(* IEC 61131-3 sources: JingjiangArm/moonboxpro_arm_8.4/Application/Application/任务列表/TensionTask/张力控制/收放料/锥度控制, 11 files *)

(* ---- StPoint_XY.st ---- *)
(*@CES
Name=StPoint_XY
Type=Gvl
TypeGuid=2db5746d-d284-4425-9f7f-2663a34b0ebc
Guid=09f53c8f-47df-4e4e-acd6-e976559a9c39
HasDeclaration=True
HasImplementation=False
*)
{DECLARATION}
TYPE StPoint_XY :(*点位置-目前用于锥度(X=卷径|Y=气压)*)
STRUCT
	rX:REAL;
	rY:REAL;
END_STRUCT
END_TYPE

{IMPLEMENTATION}

(* ---- KS_CovertUnit_Taper.st ---- *)
(*@CES
Name=KS_CovertUnit_Taper
Type=FunctionBlock
TypeGuid=6f9dac99-8de1-4efc-8465-68ac443b7d08
Guid=64151f1e-8911-4786-9206-474c18fed1e9
HasDeclaration=True
HasImplementation=True
*)
{DECLARATION}
FUNCTION KS_CovertUnit_Taper : BOOL(*锥度单位转换|以%作为基准互相转换*)
(*如果参数出错了，则会重新处理单位变量|2022.10.16.104813*)
(*2025.1.15.152522 增加了停机张力值的处理@主要时针对收料*)
VAR_INPUT
	i_pbyUnit:POINTER TO BYTE;(*单位值|0-%|1-N|2-Mpa|参数非法按照百分比显示*)
	i_xConfirmN:BOOL;(*牛顿对应确认按钮*)
	i_xConfirmMpa:BOOL;(*Mpa对应确认按钮*)
	i_prConfirmTaperPercentMatchN:POINTER TO REAL;(*确认的百分比值-牛顿单位*)
	i_prConfirmTaperPercentMatchMpa:POINTER TO REAL;(*确认的百分比值-Mpa单位*)
	i_rConfirmTaperN: REAL;(*确认的牛顿值*)
	i_rConfirmTaperMpa: REAL;(*确认的Mpa值*)
	i_prTaperValueBegin_Hmi:POINTER TO REAL;(*界面锥度显示值-起始*)
	i_prTaperValueEnd_Hmi:POINTER TO REAL;(*界面锥度显示值-结束*)
	i_prTaperValueCur_Hmi:POINTER TO REAL;(*界面显示当前值|根据单位切换*)
	i_pbyLastUnit:POINTER TO BYTE;(*上个周期的单位选择值*)

	i_prTaperPencent_Begin:POINTER TO REAL;(*锥度起始百分比值*)
	i_prTaperPencent_End:POINTER TO REAL;(*锥度起始百分比值*)
	i_lrTaperPencent_Cur:LREAL;(*锥度起始百分比当前值*)

	(*2025.1.15.152522 增加了停机张力值的处理@主要时针对收料*)
	(*不用可以写0*)
	i_pbyInitTaper:POINTER TO BYTE;(*停机初始气压百分比*)
	i_prInitTaper_Hmi:POINTER TO REAL;(*收料初始气压显示值|根据单位切换*)

END_VAR
VAR
	lrConfirmTaperPencent: LREAL;(*确认的百分比值——和*)
	lrConfirmTaper: LREAL;(*确认的百分比对应的单位的值*)

	lrCoeff: LREAL;
END_VAR
{IMPLEMENTATION}
IF i_prConfirmTaperPercentMatchN<>0 AND
	i_prConfirmTaperPercentMatchMpa<>0 AND
	i_prTaperValueBegin_Hmi<>0 AND
	i_prTaperValueEnd_Hmi<>0 AND
	i_prTaperPencent_Begin<>0 AND
	i_pbyLastUnit<>0 AND
	i_pbyUnit<>0 AND
	i_prTaperValueCur_Hmi<>0 AND
	i_prTaperPencent_End<>0 THEN;
ELSE
	RETURN;
END_IF

(*确认对应关系|*)
IF i_xConfirmN THEN(*N确认|*)
	i_prConfirmTaperPercentMatchN^:=LREAL_TO_REAL(i_lrTaperPencent_Cur);
END_IF

IF i_xConfirmMpa THEN(*Mpa确认|*)
	i_prConfirmTaperPercentMatchMpa^:=LREAL_TO_REAL(i_lrTaperPencent_Cur);
END_IF

CASE i_pbyUnit^ OF
	1:(*单位N*)
		lrConfirmTaperPencent:=i_prConfirmTaperPercentMatchN^;
		lrConfirmTaper:=i_rConfirmTaperN;

		(*2022.10.16.104832 +*)
		IF lrConfirmTaperPencent=0 OR
			lrConfirmTaper=0 THEN
			i_pbyUnit^:=0;(*确认的系数出错了|不能切换单位*)
		END_IF
	2:(*单位Mpa*)
		lrConfirmTaperPencent:=i_prConfirmTaperPercentMatchMpa^;
		lrConfirmTaper:=i_rConfirmTaperMpa;
		(*2022.10.16.104832 +*)
		IF lrConfirmTaperPencent=0 OR
			lrConfirmTaper=0 THEN
			i_pbyUnit^:=0;(*确认的系数出错了|不能切换单位*)
		END_IF
ELSE(*单位%*)
	lrConfirmTaperPencent:=0;(*根据下面条件|使用百分比显示*)
	i_pbyUnit^:=0;
END_CASE

(*单位切换了|*)
lrCoeff:=1;
IF lrConfirmTaperPencent<>0 AND  lrConfirmTaper<>0 THEN
	lrCoeff:=(lrConfirmTaper)/lrConfirmTaperPencent;
END_IF

IF i_pbyLastUnit^ <> i_pbyUnit^ THEN(*将百分比值按照对应单位换算写入*)
	i_prTaperValueBegin_Hmi^:=LREAL_TO_REAL(lrCoeff*i_prTaperPencent_Begin^);
	i_prTaperValueEnd_Hmi^:=LREAL_TO_REAL(lrCoeff*i_prTaperPencent_End^);

	(*2025.1.15.152838+针对收料起始气压的处理输出*)
	IF i_prInitTaper_Hmi<>0 AND i_pbyInitTaper<>0 THEN
		i_prInitTaper_Hmi^:=LREAL_TO_REAL(lrCoeff*i_pbyInitTaper^);
	END_IF
ELSE
	i_prTaperPencent_Begin^:=LREAL_TO_REAL(i_prTaperValueBegin_Hmi^/lrCoeff);
	i_prTaperPencent_End^:=LREAL_TO_REAL(i_prTaperValueEnd_Hmi^/lrCoeff);
	(*最大100*)
	IF i_prTaperPencent_Begin^>100 THEN i_prTaperPencent_Begin^:=100;END_IF
	IF i_prTaperPencent_End^>100 THEN i_prTaperPencent_End^:=100;END_IF

	(*2025.1.15.152838+针对收料起始气压的处理输出*)
	IF i_prInitTaper_Hmi<>0 AND i_pbyInitTaper<>0 THEN
		i_pbyInitTaper^:=LREAL_TO_BYTE(i_prInitTaper_Hmi^/lrCoeff);
		IF i_pbyInitTaper^>100 THEN i_pbyInitTaper^:=100; END_IF
	END_IF

END_IF
(*当前值根据单位转换*)
i_prTaperValueCur_Hmi^:=LREAL_TO_REAL(lrCoeff*i_lrTaperPencent_Cur);
(*更新上个周期的单位值*)
i_pbyLastUnit^:=i_pbyUnit^;

(* ---- KS_GetCurveCoeff.st ---- *)
(*@CES
Name=KS_GetCurveCoeff
Type=FunctionBlock
TypeGuid=6f9dac99-8de1-4efc-8465-68ac443b7d08
Guid=9ebd4b66-811d-4a43-a8fd-0ccbf91fd938
HasDeclaration=True
HasImplementation=True
*)
{DECLARATION}
FUNCTION KS_GetCurveCoeff : BOOL(*锥度曲线拟合系数|支持直线和二次曲线*)
(*拟合系数-直线 Y=Ax+B
	   二次曲线 Y=Ax*x+Bx+C*)

(*支持多点计算(程序中允许100点输入)*)
(*-1 参数非法
  -2 直线拟合出错了*)
VAR_INPUT
	i_byCurveType:BYTE;(*曲线类型|=0 直线
								 |=1 二次曲线(点位太少按照直线输出)
								 |=2 三次曲线(暂不支持)*)
	i_iPoitNum_Max:INT;(*最大输入的点个数|根据这个值获取点位数据*)
	i_dwSaAdr_Point_XY:DWORD;(*点位数据的首地址|按照StPoint_XY结构体存放*)
	i_piValidPoitNum:POINTER TO INT;(*最大有效点个数*)
	(*拟合系数-直线 Y=Ax+B
		   二次曲线 Y=Ax*x+Bx+C*)
	i_prFitCoeff_A:POINTER TO REAL;(*拟合系数A*)
	i_prFitCoeff_B:POINTER TO REAL;(*拟合系数B*)
	i_prFitCoeff_C:POINTER TO REAL;(*拟合系数C*)
END_VAR
VAR
	in: INT;
	iPoitNum_Max: INT;(*最大点数*)
	astStPoint_XY:ARRAY [1..100] OF StPoint_XY;(*X轴为卷径|Y 为锥度值@按照100个点申请*)
	astValidStPoint_XY:ARRAY [1..100] OF StPoint_XY;(*X轴为卷径|Y 为锥度值@有效的点位*)
	iValidPoitNum:INT;(*有效点位的个数*)
	byCurveType: BYTE;(*曲线类型*)
	rA: REAL;
	rB: REAL;
	rC: REAL;
	xRtn: BOOL;
	iErrCode:INT;
END_VAR
{IMPLEMENTATION}
byCurveType:=i_byCurveType;
iPoitNum_Max:=i_iPoitNum_Max;
IF i_dwSaAdr_Point_XY<>0 THEN;
	SysMemCpy(ADR(astStPoint_XY),i_dwSaAdr_Point_XY,INT_TO_DWORD(iPoitNum_Max)*SIZEOF(astStPoint_XY[1]));
ELSE
	iErrCode:=-1;
END_IF

(*检查点位的合法性-X或者Y有一个=0认为是无效点*)
FOR iN:=1 TO iPoitNum_Max BY 1 DO
	IF astStPoint_XY[iN].rX=0 OR
		astStPoint_XY[iN].rY=0 THEN(*非法点，剔除*);
	ELSE
		iValidPoitNum:=iValidPoitNum+1;
		astValidStPoint_XY[iValidPoitNum]:=astStPoint_XY[iN];
	END_IF
END_FOR

(*曲线算法*)
byCurveType:=i_byCurveType;
CASE byCurveType OF
	0:(*直线拟合|*)
		xRtn:=KS_StraightLine(iValidPoitNum, ADR(astValidStPoint_XY), ADR(rA), ADR(rB));
		IF xRtn THEN
			iErrCode:=-2;
		END_IF
ELSE(*默认按照二次拟合*)
		xRtn:=KS_ParabolicLine(
					iValidPoitNum(*i_iValidPoitNum*),
					ADR(astValidStPoint_XY)(*i_pastValidStPoint_XY*),
					ADR(rA)(*i_prA*),
					ADR(rB)(*i_prB*),
					ADR(rC)(*i_prC*));
		IF xRtn THEN
			iErrCode:=-2;
		END_IF
END_CASE

IF i_piValidPoitNum<>0 THEN
	i_piValidPoitNum^:=iValidPoitNum;
END_IF
IF i_prFitCoeff_A<>0 THEN
	i_prFitCoeff_A^:=rA;
END_IF
IF i_prFitCoeff_B<>0 THEN
	i_prFitCoeff_B^:=rB;
END_IF

IF i_prFitCoeff_C<>0 THEN
	i_prFitCoeff_C^:=rC;
END_IF

KS_GetCurveCoeff:=iErrCode<>0;

(* ---- KS_ParabolicLine.st ---- *)
(*@CES
Name=KS_ParabolicLine
Type=FunctionBlock
TypeGuid=6f9dac99-8de1-4efc-8465-68ac443b7d08
Guid=32bb2783-1164-4a85-bd37-5e8616daa227
HasDeclaration=True
HasImplementation=True
*)
{DECLARATION}
FUNCTION KS_ParabolicLine : BOOL(*二次抛物线|Y=Ax^2+Bx+C@先不处理多点直线拟合|输出有效则报错*)
VAR_INPUT
	i_iValidPoitNum:INT;(*最大有效点个数*)
	i_pastValidStPoint_XY:POINTER TO ARRAY [1..100] OF StPoint_XY;(*X轴为卷径|Y 为锥度值@有效的点位*)
	i_prA:POINTER TO REAL;
	i_prB:POINTER TO REAL;
	i_prC:POINTER TO REAL;
END_VAR
VAR
	xParaErr:BOOL;
	arPoint_X:ARRAY [1..100] OF REAL;
	arPoint_Y:ARRAY [1..100] OF REAL;
	lrATemp:LREAL;
	lrBTemp:LREAL;
	rA:REAL;
	rB:REAL;
	rC:REAL;
	iN: INT;
	byType: BYTE;
	pstValidStPoint_XY:POINTER TO StPoint_XY;(*X轴为卷径|Y 为锥度值@有效的点位*)
	lrTemp: LREAL;
	lrTemp1: LREAL;
	lrTemp2: LREAL;
	lrTemp3: LREAL;
	lrTemp4: LREAL;
	lrTemp5: LREAL;
	lrTemp6: LREAL;
	lrTemp7: LREAL;
	lrAverage_X: LREAL;(*X的平均值*)
	lrAverage_Y: LREAL;(*Y的平均值*)
	lrAverage_XY: LREAL;(*XY的平均值*)
	lrAverage_X_Square2: LREAL;(*X^2的平均值*)
	lrAverage_X_Square3: LREAL;(*X^3的平均值*)
	lrAverage_X_Square4: LREAL;(*X^4的平均值*)
	lrAverage_XSquare2Y: LREAL;(*X^2*Y的平均值*)
END_VAR
{IMPLEMENTATION}
IF i_pastValidStPoint_XY<>0 THEN
	IF i_iValidPoitNum>=4 THEN(*4个点以上使用拟合算法*)
		byType:=3;
	ELSIF i_iValidPoitNum=3 THEN(*3个点使用抛物线*)
		byType:=2;
	ELSIF i_iValidPoitNum=2 THEN(*2个点使用直线*)
		byType:=1;
	ELSE(*点位太少*)
		xParaErr:=TRUE;
	END_IF

	IF NOT xParaErr THEN
		FOR iN:=1  TO i_iValidPoitNum BY 1 DO
			pstValidStPoint_XY:=ADR(i_pastValidStPoint_XY^[iN]);
			arPoint_X[iN]:=pstValidStPoint_XY^.rX;
			arPoint_Y[iN]:=pstValidStPoint_XY^.rY;
		END_FOR

		CASE byType OF
			1:(*直线*)
				lrTemp	:=arPoint_X[1]-arPoint_X[2];
				lrTemp1	:=arPoint_Y[1]-arPoint_Y[2];
				IF lrTemp<>0 THEN
					rA:=LREAL_TO_REAL(lrTemp1/lrTemp);

					lrTemp1:=arPoint_X[1]*arPoint_Y[2]-arPoint_X[2]*arPoint_Y[1];
					rB:=lrTemp1/lrTemp;
				ELSE
					xParaErr:=TRUE;
				END_IF

			2:(*抛物线*)
				(*计算rB*)
				lrTemp1:=(arPoint_X[2]*arPoint_X[2]-arPoint_X[3]*arPoint_X[3]);(*X2^2-X3^2*)
				lrTemp1:=lrTemp1*(arPoint_X[1]-arPoint_X[2]);(*lrTemp1*(X1-X2)*)
				lrTemp2:=(arPoint_X[1]*arPoint_X[1]-arPoint_X[2]*arPoint_X[2]);(*X1^2-X2^2*)
				lrTemp2:=lrTemp2*(arPoint_X[2]-arPoint_X[3]);(*lrTemp2*(X2-X3)*)
				lrTemp:=lrTemp1-lrTemp2;(*rB的分母*)

				IF lrTemp<>0 THEN
					lrTemp1:=(arPoint_X[2]*arPoint_X[2]-arPoint_X[3]*arPoint_X[3]);(*X2^2-X3^2*)
					lrTemp1:=lrTemp1*(arPoint_Y[1]-arPoint_Y[2]);(*lrTemp1*(Y1-Y2)*)
					lrTemp2:=(arPoint_X[1]*arPoint_X[1]-arPoint_X[2]*arPoint_X[2]);(*X1^2-X2^2*)
					lrTemp2:=lrTemp2*(arPoint_Y[2]-arPoint_Y[3]);(*lrTemp1*(Y2-Y3)*)

					rB:=(lrTemp1-lrTemp2)/lrTemp;
				ELSE
					xParaErr:=TRUE;
				END_IF

				(*计算rA*)
				IF NOT xParaErr THEN
					lrTemp:=(arPoint_X[1]*arPoint_X[1]-arPoint_X[2]*arPoint_X[2]);(*X1^2-X2^2*)
					IF lrTemp<>0 THEN
						lrTemp1:=arPoint_Y[1]-arPoint_Y[2]-rB*(arPoint_X[1]-arPoint_X[2]);(*Y1-Y2-rB*(X1-X2)*)
						rA:=lrTemp1/lrTemp;
					ELSE
						xParaErr:=TRUE;
					END_IF
				END_IF
				(*计算rC*)
				IF NOT xParaErr THEN
					rC:=arPoint_Y[1]-rA*(arPoint_X[1]*arPoint_X[1])-rB*arPoint_X[1];
				END_IF

			3:(*拟合曲线|*)
				lrTemp:=0;
				lrTemp1:=0;
				lrTemp2:=0;
				lrTemp3:=0;
				lrTemp4:=0;
				lrTemp5:=0;
				lrTemp6:=0;
				lrTemp7:=0;
				FOR iN:=1 TO i_iValidPoitNum BY 1 DO
					lrTemp1:=lrTemp1+arPoint_X[iN];
					lrTemp2:=lrTemp2+arPoint_Y[iN];
					lrTemp3:=lrTemp3+arPoint_X[iN]*arPoint_Y[iN];
					lrTemp4:=lrTemp4+arPoint_X[iN]*arPoint_X[iN];
					lrTemp5:=lrTemp5+arPoint_X[iN]*arPoint_X[iN]*arPoint_X[iN];
					lrTemp6:=lrTemp6+arPoint_X[iN]*arPoint_X[iN]*arPoint_X[iN]*arPoint_X[iN];
					lrTemp7:=lrTemp7+arPoint_X[iN]*arPoint_X[iN]*arPoint_Y[iN];
				END_FOR

				(*计算X Y的平均值*)
				lrAverage_X			:=lrTemp1/i_iValidPoitNum;
				lrAverage_Y			:=lrTemp2/i_iValidPoitNum;
				lrAverage_XY		:=lrTemp3/i_iValidPoitNum;
				lrAverage_X_Square2	:=lrTemp4/i_iValidPoitNum;
				lrAverage_X_Square3	:=lrTemp5/i_iValidPoitNum;
				lrAverage_X_Square4	:=lrTemp6/i_iValidPoitNum;
				lrAverage_XSquare2Y	:=lrTemp7/i_iValidPoitNum;

				(*计算拟合的rA*)
				lrTemp1:=lrAverage_X_Square3-lrAverage_X*lrAverage_X_Square2;
				lrTemp1:=lrTemp1*lrTemp1;
				lrTemp2:=lrAverage_X_Square4-lrAverage_X_Square2*lrAverage_X_Square2;
				lrTemp2:=lrTemp2*(lrAverage_X_Square2-lrAverage_X*lrAverage_X);
				lrTemp:=lrTemp1-lrTemp2;(*计算分母*)
				IF lrTemp<>0 THEN
					lrTemp1:=lrAverage_XY-lrAverage_X*lrAverage_Y;
					lrTemp1:=lrTemp1*(lrAverage_X_Square3-lrAverage_X*lrAverage_X_Square2);

					lrTemp2:=lrAverage_XSquare2Y-lrAverage_X_Square2*lrAverage_Y;
					lrTemp2:=lrTemp2*(lrAverage_X_Square2-lrAverage_X*lrAverage_X);
					lrATemp:=(lrTemp1-lrTemp2)/lrTemp;
					rA:=lrATemp;
				ELSE
					xParaErr:=TRUE;
				END_IF
				(*计算rB*)
				IF NOT xParaErr THEN
					lrTemp:=lrAverage_X_Square2-lrAverage_X*lrAverage_X;
					IF lrTemp<>0 THEN
						lrTemp1:=lrAverage_XY-lrAverage_X*lrAverage_Y-lrATemp*(lrAverage_X_Square3-lrAverage_X*lrAverage_X_Square2);
						lrBTemp:=lrTemp1/lrTemp;
						rB:=lrBTemp;
					ELSE
						xParaErr:=TRUE;
					END_IF
				END_IF

				(*计算rC*)
				IF NOT xParaErr THEN
					lrTemp:=lrAverage_Y-lrATemp*lrAverage_X_Square2-lrBTemp*lrAverage_X;
					rC:=lrTemp;
				END_IF
		ELSE;
		END_CASE

	END_IF
ELSE
	xParaErr:=TRUE;
END_IF

IF i_prA<>0 THEN
	i_prA^:=rA;
END_IF

IF i_prB<>0 THEN
	i_prB^:=rB;
END_IF

IF i_prC<>0 THEN
	i_prC^:=rC;
END_IF

KS_ParabolicLine:=xParaErr;

(* ---- KS_StraightLine.st ---- *)
(*@CES
Name=KS_StraightLine
Type=FunctionBlock
TypeGuid=6f9dac99-8de1-4efc-8465-68ac443b7d08
Guid=69642510-d218-426d-a290-8472573a37ba
HasDeclaration=True
HasImplementation=True
*)
{DECLARATION}
FUNCTION KS_StraightLine : BOOL(*直线|Y=Ax+B@先不处理多点直线拟合|输出有效则报错*)
VAR_INPUT
	i_iValidPoitNum:INT;(*最大有效点个数*)
	i_pastValidStPoint_XY:POINTER TO ARRAY [1..100] OF StPoint_XY;(*X轴为卷径|Y 为锥度值@有效的点位*)
	i_prA:POINTER TO REAL;
	i_prB:POINTER TO REAL;
END_VAR
VAR
	xParaErr:BOOL;
	arPoint_X:ARRAY [1..100] OF REAL;
	arPoint_Y:ARRAY [1..100] OF REAL;
	rA:REAL;
	rB:REAL;
	iN: INT;
	byType: BYTE;
	pstValidStPoint_XY:POINTER TO StPoint_XY;(*X轴为卷径|Y 为锥度值@有效的点位*)
	lrTemp: LREAL;
	lrTemp1: LREAL;
	lrTemp2: LREAL;
	lrTemp3: LREAL;
	lrTemp4: LREAL;
	lrSum_X: LREAL;
	lrSum_Y: LREAL;
	lrSum_XY: LREAL;
	lrSum_XSquart2: LREAL;
END_VAR
{IMPLEMENTATION}
IF i_pastValidStPoint_XY<>0 THEN
	IF i_iValidPoitNum>=3 THEN(*3个点以上使用拟合算法*)
		byType:=2;
	ELSIF i_iValidPoitNum=2 THEN(*2个点使用直线*)
		byType:=1;
	ELSE(*点位太少*)
		xParaErr:=TRUE;
	END_IF

	IF NOT xParaErr THEN
		FOR iN:=1  TO i_iValidPoitNum BY 1 DO
			pstValidStPoint_XY:=ADR(i_pastValidStPoint_XY^[iN]);
			arPoint_X[iN]:=pstValidStPoint_XY^.rX;
			arPoint_Y[iN]:=pstValidStPoint_XY^.rY;
		END_FOR

		CASE byType OF
			1:(*直线*)
				lrTemp	:=arPoint_X[1]-arPoint_X[2];
				lrTemp1	:=arPoint_Y[1]-arPoint_Y[2];
				IF lrTemp<>0 THEN
					rA:=LREAL_TO_REAL(lrTemp1/lrTemp);

					lrTemp1:=arPoint_X[1]*arPoint_Y[2]-arPoint_X[2]*arPoint_Y[1];
					rB:=LREAL_TO_REAL(lrTemp1/lrTemp);
				ELSE
					xParaErr:=TRUE;
				END_IF

			2:(*拟合直线*)
				lrSum_X:=0;
				lrSum_Y:=0;
				lrSum_XY:=0;
				lrSum_XSquart2:=0;
				FOR iN:=1 TO i_iValidPoitNum BY 1 DO
					lrSum_X:=lrSum_X+arPoint_X[iN];
					lrSum_Y:=lrSum_Y+arPoint_Y[iN];
					lrSum_XY:=lrSum_XY+arPoint_X[iN]*arPoint_Y[iN];
					lrSum_XSquart2:=lrSum_XSquart2+arPoint_X[iN]*arPoint_X[iN];
				END_FOR

				(*计算rB*)
				lrTemp:=i_iValidPoitNum*lrSum_XSquart2-lrSum_X*lrSum_X;
				IF lrTemp<>0 THEN
					lrTemp1:=lrSum_XSquart2*lrSum_Y-lrSum_X*lrSum_XY;
					rB:=LREAL_TO_REAL(lrTemp1/lrTemp);
				ELSE
					xParaErr:=TRUE;
				END_IF

				(*计算rA*)
				IF NOT xParaErr THEN
					lrTemp:=i_iValidPoitNum*lrSum_XSquart2-lrSum_X*lrSum_X;
					IF lrTemp<>0 THEN
						lrTemp1:=i_iValidPoitNum*lrSum_XY-lrSum_X*lrSum_Y;
						rA:=LREAL_TO_REAL(lrTemp1/lrTemp);
					ELSE
						xParaErr:=TRUE;
					END_IF
				END_IF
		ELSE;
		END_CASE

	END_IF
ELSE
	xParaErr:=TRUE;
END_IF

IF i_prA<>0 THEN
	i_prA^:=rA;
END_IF

IF i_prB<>0 THEN
	i_prB^:=rB;
END_IF

KS_StraightLine:=xParaErr;

(* ---- KS_Taper_Curve.st ---- *)
(*@CES
Name=KS_Taper_Curve
Type=FunctionBlock
TypeGuid=6f9dac99-8de1-4efc-8465-68ac443b7d08
Guid=9d8a75d4-e332-49bf-ad4d-ef60c80700c3
HasDeclaration=True
HasImplementation=True
*)
{DECLARATION}
FUNCTION KS_Taper_Curve : LREAL(*锥度1/X算法*)(*输出当前锥度*)
(*2025.1.9.162727  增加当前卷径输入*)
(*2025.2.26.163100 bug处理*)
VAR_INPUT
	i_rDiamCurAxis_Rw:REAL;(*2025.1.9.162744+*)
	i_rTaper_Begin_Rw: REAL;(*起始锥度*)
	i_rTaper_End_Rw: REAL;(*结束锥度*)
	i_rDiamTaper_Begin_Rw: REAL;(*起始锥度-直径*)
	i_rDiamTaper_End_Rw: REAL;(*结束锥度-直径*)
END_VAR
VAR
	lrMomentSa: LREAL;(*起始力矩*)
	lrMomentEd: LREAL;(*结束力矩*)
	lrCurrentMoment: LREAL;(*当前力矩*)
	lrCurrentTaper:LREAL;
END_VAR
{IMPLEMENTATION}
lrCurrentTaper:=0;
lrMomentSa:=(i_rTaper_Begin_Rw)*i_rDiamTaper_Begin_Rw;
lrMomentEd:=(i_rTaper_End_Rw)*i_rDiamTaper_End_Rw;

(*取消该限制@2025.2.26.163020*)
(*	IF lrMomentEd< lrMomentSa THEN lrMomentEd:=lrMomentSa;END_IF*)

IF i_rDiamCurAxis_Rw<= i_rDiamTaper_Begin_Rw THEN
	(*最小卷用最大张力*)
	lrCurrentTaper:= i_rTaper_Begin_Rw;
ELSIF i_rDiamCurAxis_Rw>= i_rDiamTaper_End_Rw THEN
	(*最大卷用最小张力*)
	lrCurrentTaper:= i_rTaper_End_Rw;
ELSE
	IF ( i_rDiamTaper_End_Rw-i_rDiamTaper_Begin_Rw)<>0 THEN
		lrCurrentMoment:=lrMomentSa+(lrMomentEd-lrMomentSa)*(i_rDiamCurAxis_Rw-i_rDiamTaper_Begin_Rw)
						/(i_rDiamTaper_End_Rw-i_rDiamTaper_Begin_Rw);
	ELSE
		lrCurrentMoment:=lrMomentSa;
	END_IF

	IF i_rDiamCurAxis_Rw<>0 THEN
		lrCurrentTaper:=lrCurrentMoment/i_rDiamCurAxis_Rw;
	ELSE
		lrCurrentTaper:=i_rTaper_Begin_Rw;
	END_IF
END_IF

KS_Taper_Curve:=lrCurrentTaper;

(* ---- KS_Taper_Straight.st ---- *)
(*@CES
Name=KS_Taper_Straight
Type=FunctionBlock
TypeGuid=6f9dac99-8de1-4efc-8465-68ac443b7d08
Guid=74716efb-2a9a-4cd3-af40-131a820a6ef5
HasDeclaration=True
HasImplementation=True
*)
{DECLARATION}
FUNCTION KS_Taper_Straight : LREAL(*锥度直线算法*)(*输出当前锥度*)
(*2025.1.9.162837 增加当前卷径输入*)
VAR_INPUT
	i_rDiamCurAxis_Rw:REAL;
	i_rTaper_Begin_Rw: REAL;(*起始锥度*)
	i_rTaper_End_Rw: REAL;(*结束锥度*)
	i_rDiamTaper_Begin_Rw: REAL;(*起始锥度-直径*)
	i_rDiamTaper_End_Rw: REAL;(*结束锥度-直径*)
END_VAR
VAR
	lrTempPercent: LREAL; (*临时用来计算%的变量*)
	lrCurrentTaper:LREAL;
END_VAR
{IMPLEMENTATION}
lrCurrentTaper:=0;
IF i_rDiamTaper_Begin_Rw<i_rDiamTaper_End_Rw THEN
	IF i_rDiamCurAxis_Rw<=i_rDiamTaper_Begin_Rw THEN
		(*最小卷用最大张力*)
		lrCurrentTaper:= i_rTaper_Begin_Rw;
	ELSIF i_rDiamCurAxis_Rw>=i_rDiamTaper_End_Rw THEN
		(*最大卷用最小张力*)
		lrCurrentTaper:= i_rTaper_End_Rw;
	ELSE
		(*卷径锥度的线性关系有效*)
		lrTempPercent:= (i_rDiamCurAxis_Rw - i_rDiamTaper_Begin_Rw) / (i_rDiamTaper_End_Rw - i_rDiamTaper_Begin_Rw);
		lrCurrentTaper:= i_rTaper_Begin_Rw - lrTempPercent * (i_rTaper_Begin_Rw - i_rTaper_End_Rw);
	END_IF
ELSE
	lrCurrentTaper:= 0;
END_IF
KS_Taper_Straight:=lrCurrentTaper;

(* ---- KS_FB_Taper.st ---- *)
(*@CES
Name=KS_FB_Taper
Type=FunctionBlock
TypeGuid=6f9dac99-8de1-4efc-8465-68ac443b7d08
Guid=684df15a-86b3-4c73-bdbe-f6eb8637542a
HasDeclaration=True
HasImplementation=True
*)
{DECLARATION}
FUNCTION_BLOCK KS_FB_Taper
(*2025.1.9.162926 增加了当前卷径输入接口@写到输入输出是为了防止漏改*)
(*2025.1.15.150823 停机锥度@防止停机张力投入时收料锥度设置过小引起的料膜被放料拉走问题*)
(*2025.3.7.112920 增加了多点直线和多点曲线的实现*)
(*2025.3.29.151033 停机锥度的实现更新丢了！麻烦*)
VAR_INPUT
	i_iGrpId: INT; (*1.A系;2.B系*)
	i_xTaperCurCTLEn:BOOL;(*当前锥度控制使能|在印刷状态且收牵合压或者色组至少合压一色时进行控制
						其他状态按照最大锥度输出|2021.8.30.164822*)
//	i_pstStShmGlobalParam: POINTER TO StShmGlobalParam; (*参数地址*)
	i_xTaperAdd:BOOL;
	i_xTaperDec:BOOL;
	i_rTaperMax:REAL;(*最大锥度限值值*)
	i_rTaperValue_Stop:REAL;(*停机锥度@防止停机张力投入时收料锥度设置过小引起的料膜被放料拉走问题*)

	i_byTaperAdjMode: BYTE;
	i_rDiamCurAxis: REAL;
	i_rTaper_Begin_Rw: REAL;(*起始锥度*)
	i_rTaper_End_Rw: REAL;(*结束锥度*)
	i_rDiamTaper_Begin_Rw: REAL;(*起始锥度-直径*)
	i_rDiamTaper_End_Rw: REAL;(*结束锥度-直径*)
END_VAR
VAR_OUTPUT
	o_rTaper_Cur: REAL;
END_VAR
VAR_IN_OUT
	iO_byTaperUnit: BYTE;
	io_rTaperValueBegin_Hmi: REAL;
	io_rTaperValueEnd_Hmi: REAL;
	io_astTaperPoint:ARRAY [1..10] OF StPoint_XY;
END_VAR
VAR
//	pstStGrpParam: POINTER TO StGrpParam; (*访问当前系参数的指针*)
	xTaperAdd:BOOL;
	xPreTaperAdd:BOOL;
	xTaperDec:BOOL;
	xPreTaperDec:BOOL;
	lrTemp: LREAL;
	lrCurrentTaper: LREAL;(*当前锥度值临时变量*)

	lrPreCurrentTaper: LREAL;(*上个周期的锥度*)
	lrDelTaper: LREAL;(*锥度的变化量*)
	iMaxTimeTOMaxTaper:INT:=200;(*到达最大锥度的周期次数，20ms周期时时间是4s*)
	iMaxTaper:INT:=100;(*最大锥度值*)

	(*2025.3.7.113256+byTaperAdjMode = 2*)
	xRtn: BOOL;
	iN: INT;
	iPoitMax: INT:=7;(*最大点数先按照7个*)
	iValidPoitNum: INT;(*实际有效的点数*)
	rFitCoeff_A: REAL;(*计算的二次系数*)
	rFitCoeff_B: REAL;(*计算的一次系数*)
	rFitCoeff_C: REAL;(*常量*)
	iMaxDiamIndex: INT;(*多点中卷径最大值索引*)
	iMinDiamIndex: INT;(*多点中卷径最小值索引*)
	rMinDiam: REAL;(*多点中最小卷径值*)
	rMaxDiam: REAL;(*多点中最大卷径值*)
END_VAR
{IMPLEMENTATION}
IF (i_iGrpId=1 OR i_iGrpId=2) THEN ;ELSE RETURN;END_IF

//pstStGrpParam:= ADR(i_pstStShmGlobalParam^.astStGrpParam[i_iGrpId]);

xTaperAdd:= i_xTaperAdd;
xTaperDec:= i_xTaperDec;

(*2022.2.23.112107 调整锥度界面加减逻辑*)
IF iO_byTaperUnit=1 THEN(*单位是N*)
	lrTemp:=1;
ELSIF iO_byTaperUnit=2 THEN(*单位是mpa*)
	lrTemp:=0.01;
ELSE(*单位是%*)
	lrTemp:=1;
END_IF

IF xTaperAdd AND NOT xPreTaperAdd THEN
	lrTemp:=lrTemp;
ELSIF xTaperDec AND NOT xPreTaperDec THEN
	lrTemp:=-lrTemp;
ELSE
	lrTemp:=0;
END_IF
(*
pstStGrpParam^.lrTaper_Begin_Rw:= pstStGrpParam^.lrTaper_Begin_Rw+lrTemp;
pstStGrpParam^.lrTaper_End_Rw:= pstStGrpParam^.lrTaper_End_Rw+lrTemp;
*)
(*2022.2.23.112206 处理的变量修改为带hmi界面的*)

io_rTaperValueBegin_Hmi:= io_rTaperValueBegin_Hmi+lrTemp;
io_rTaperValueEnd_Hmi:= io_rTaperValueEnd_Hmi+lrTemp;

IF 	io_rTaperValueBegin_Hmi>i_rTaperMax THEN
	io_rTaperValueBegin_Hmi:= i_rTaperMax;
ELSIF io_rTaperValueBegin_Hmi<0 THEN
	io_rTaperValueBegin_Hmi:=0;
END_IF

IF 	io_rTaperValueEnd_Hmi>i_rTaperMax THEN
	io_rTaperValueEnd_Hmi:= i_rTaperMax;
ELSIF io_rTaperValueEnd_Hmi<0 THEN
	io_rTaperValueEnd_Hmi:=0;
END_IF

xPreTaperAdd:=xTaperAdd;
xPreTaperDec:=xTaperDec;

(*
(*2019.4.11.164149 将锥度控制移植到功能块中.并额外增加了新的算法*)
CASE i_pstStShmGlobalParam^.stStSystemExtInfo.byTaperAdjMode OF
1:
	lrCurrentTaper:=KS_Taper_Curve(pstStGrpParam^.lrDiamCurAxis_Rw,pstStGrpParam);
ELSE
	lrCurrentTaper:=KS_Taper_Straight(pstStGrpParam^.lrDiamCurAxis_Rw,pstStGrpParam);
END_CASE

(*2021.8.30.164530 |*)
(*不控制的时候按照最大锥度输出*)
IF NOT i_xTaperCurCTLEn THEN
	lrCurrentTaper:=MAX(pstStGrpParam^.lrTaper_Begin_Rw,pstStGrpParam^.lrTaper_End_Rw);(*取最大值*)
	(*增加一个变量单独控制停机的锥度*)
	lrCurrentTaper:=MAX(lrCurrentTaper,i_rTaperValue_Stop);
END_IF
*)

(*2025.3.7.112958 +*)
(*2019.4.11.164149 将锥度控制移植到功能块中.并额外增加了新的算法*)
(*0--2变化*)
xRtn:=FALSE;
CASE i_byTaperAdjMode OF
1:(*2点曲线*)

	lrCurrentTaper:=KS_Taper_Curve(
			i_rDiamCurAxis,
			i_rTaper_Begin_Rw,
			i_rTaper_End_Rw,
			i_rDiamTaper_Begin_Rw,
			i_rDiamTaper_End_Rw
			);

	(*2021.8.30.164530 |*)
	(*不控制的时候按照最大锥度输出*)
	IF NOT i_xTaperCurCTLEn THEN
(*
		lrCurrentTaper:=MAX(pstStGrpParam^.lrTaper_Begin_Rw,pstStGrpParam^.lrTaper_End_Rw);(*取最大值*)
		(*增加一个变量单独控制停机的锥度*)
		lrCurrentTaper:=MAX(lrCurrentTaper,i_rTaperValue_Stop);
*)
		(*2025.3.29.151947+*)
		lrCurrentTaper:=i_rTaperValue_Stop;
	END_IF

2:(*多点曲线@2025.2.28.235627+*)
	(*寻找卷径锥度的最大值和最小值@限制输出使用*)
	iMinDiamIndex:=0;
	iMaxDiamIndex:=0;
	FOR iN:=1 TO iPoitMax BY 1 DO
		(*最小卷径值的索引*)
		IF iMinDiamIndex=0 THEN(*先找起始索引*)
			IF io_astTaperPoint[iN].rX<>0 THEN
				iMinDiamIndex:=iN;
			END_IF
		ELSE(*找到了第一个值*)
			IF io_astTaperPoint[iN].rX < io_astTaperPoint[iMinDiamIndex].rX THEN
				iMinDiamIndex:=iN;(*更新索引值*)
			END_IF
		END_IF

		(*最大卷径的索引*)
		IF iMaxDiamIndex=0 THEN(*先找起始索引*)
			IF io_astTaperPoint[iN].rX<>0 THEN
				iMaxDiamIndex:=iN;
			END_IF
		ELSE(*找到了第一个值*)
			IF io_astTaperPoint[iN].rX > io_astTaperPoint[iMaxDiamIndex].rX THEN
				iMaxDiamIndex:=iN;(*更新索引值*)
			END_IF
		END_IF
	END_FOR

	xRtn:=KS_GetCurveCoeff(
			1(*i_byCurveType*),
			iPoitMax(*i_iPoitNum_Max*),
			ADR(io_astTaperPoint[1])(*i_dwSaAdr_Point_XY*),
			ADR(iValidPoitNum)(*i_piValidPoitNum*),
			ADR(rFitCoeff_A)(*i_prFitCoeff_A*),
			ADR(rFitCoeff_B)(*i_prFitCoeff_B*),
			ADR(rFitCoeff_C)(*i_prFitCoeff_C*));
	(*输出的形式是a*x*x+b*x+C*)
	IF NOT xRtn THEN(*未报错@至少2个点*)
		lrCurrentTaper:=rFitCoeff_A*i_rDiamCurAxis*i_rDiamCurAxis+
						rFitCoeff_B*i_rDiamCurAxis+
						rFitCoeff_C;
		(*限值处理*)
		IF	iMinDiamIndex>0 AND iMinDiamIndex<=iPoitMax AND(*索引合法判断*)
			iMaxDiamIndex>0 AND iMaxDiamIndex<=iPoitMax THEN(*索引合法判断*)
			(*最小值处理*)
			rMinDiam:= io_astTaperPoint[iMinDiamIndex].rX;
			IF i_rDiamCurAxis<=rMinDiam THEN
				lrCurrentTaper:=rFitCoeff_A*rMinDiam*rMinDiam+
								rFitCoeff_B*rMinDiam+
								rFitCoeff_C;
			END_IF
			(*最大值处理*)
			rMaxDiam:= io_astTaperPoint[iMaxDiamIndex].rX;
			IF i_rDiamCurAxis>=rMaxDiam THEN
				lrCurrentTaper:=rFitCoeff_A*rMaxDiam*rMaxDiam+
								rFitCoeff_B*rMaxDiam+
								rFitCoeff_C;
			END_IF
(*
			(*2025.3.3.112928 调整*)
			(*2021.8.30.164530 |*)
			(*不控制的时候按照最大锥度输出*)
			IF NOT i_xTaperCurCTLEn THEN
				lrCurrentTaper:=MAX(rFitCoeff_A*rMinDiam*rMinDiam+rFitCoeff_B*rMinDiam+rFitCoeff_C,
								rFitCoeff_A*rMaxDiam*rMaxDiam+rFitCoeff_B*rMaxDiam+rFitCoeff_C);(*取最大值*)
				(*增加一个变量单独控制停机的锥度*)
				lrCurrentTaper:=MAX(lrCurrentTaper,i_rTaperValue_Stop);

			END_IF
*)
		ELSE
			lrCurrentTaper:=22.2;(*就随便给一个特殊值吧@有可能能指导查找问题*)
		END_IF
	ELSE(*拟合失败了@按照最大点输出*)
		IF iMaxDiamIndex>0 AND iMaxDiamIndex<=iPoitMax THEN(*索引合法判断*)
			lrCurrentTaper:=io_astTaperPoint[iMaxDiamIndex].rY;
		END_IF
	END_IF

	(*2025.3.29.151918+*)
	(*不控制的时候按照最大锥度输出*)
	IF NOT i_xTaperCurCTLEn THEN
		lrCurrentTaper:=i_rTaperValue_Stop;
	END_IF
ELSE(*2点直线*)
	lrCurrentTaper:=KS_Taper_Straight(
			i_rDiamCurAxis,
			i_rTaper_Begin_Rw,
			i_rTaper_End_Rw,
			i_rDiamTaper_Begin_Rw,
			i_rDiamTaper_End_Rw
			);

	(*2021.8.30.164530 |*)
	(*不控制的时候按照最大锥度输出*)
	IF NOT i_xTaperCurCTLEn THEN
(*
		lrCurrentTaper:=MAX(pstStGrpParam^.lrTaper_Begin_Rw,pstStGrpParam^.lrTaper_End_Rw);(*取最大值*)
		(*增加一个变量单独控制停机的锥度*)
		lrCurrentTaper:=MAX(lrCurrentTaper,i_rTaperValue_Stop);
*)
		(*2025.3.29.151937+*)
		lrCurrentTaper:=i_rTaperValue_Stop;
	END_IF
END_CASE

lrDelTaper:=INT_TO_LREAL(iMaxTaper)/INT_TO_LREAL(iMaxTimeTOMaxTaper);
(*rWatch:=lrCurrentTaper;*)
IF lrCurrentTaper> lrPreCurrentTaper THEN
	IF (lrCurrentTaper-lrPreCurrentTaper) > lrDelTaper THEN
		lrCurrentTaper:=lrPreCurrentTaper+lrDelTaper;
	ELSE;
	END_IF
ELSIF  lrCurrentTaper< lrPreCurrentTaper THEN
	IF (lrPreCurrentTaper-lrCurrentTaper) > lrDelTaper THEN
		lrCurrentTaper:=lrPreCurrentTaper-lrDelTaper;
	ELSE;
	END_IF
ELSE;
END_IF

o_rTaper_Cur:= LREAL_TO_REAL(lrCurrentTaper);
lrPreCurrentTaper:=lrCurrentTaper;

(* ---- KS_FB_Taper_UwRw_IfOf.st ---- *)
(*@CES
Name=KS_FB_Taper_UwRw_IfOf
Type=FunctionBlock
TypeGuid=6f9dac99-8de1-4efc-8465-68ac443b7d08
Guid=4508f757-99f8-49ac-966d-1f120aaadfc2
HasDeclaration=True
HasImplementation=True
*)
{DECLARATION}
FUNCTION_BLOCK KS_FB_Taper_UwRw_IfOf
VAR_INPUT
	i_xEn: BOOL;
END_VAR
VAR_OUTPUT
END_VAR
VAR
	fbKS_FB_TaperUnitDeal: KS_FB_TaperUnitDeal;
	(*锥度变化临时变量|只处理放料 放牵收牵*)
	rMaxTaper:REAL:=100;(*最大锥度|目前使用%*)
	iTimeTaperChange:INT:=10000;(*锥度变化时间|ms*)
	rTaperTar: REAL;
	rTaperCur: REAL;
	rDeltTaper: REAL;
	xInit_Taper_Cur: BOOL;
END_VAR
{IMPLEMENTATION}
IF i_xEn THEN
	(*2021.7.29.094016 张力单位切换控制逻辑|以及标定逻辑*)
	fbKS_FB_TaperUnitDeal(i_pstStGrpParam:=pstStGrpParam );

	(*处理4个锥度|放料、放牵、收料、收牵*)
	(*需要确定是否需要进行单位转换|目前是%*)
	(*使用起始锥度作为界面显示|当前锥度做规划*)
	(*放料*)
	(*由于当前锥度是保持型的|在这里做开机初始复位处理|*)
	IF NOT xInit_Taper_Cur THEN
		xInit_Taper_Cur:=TRUE;
		pstStGrpParam^.lrTaper_Cur_Uw:=0;
		pstStGrpParam^.lrTaper_Cur_If:=0;
		pstStGrpParam^.lrTaper_Cur_Of:=0;
	END_IF

	rTaperTar:=pstStGrpParam^.lrTaper_Begin_Uw;
	rTaperCur:=pstStGrpParam^.lrTaper_Cur_Uw;
	rDeltTaper:=rMaxTaper/iTimeTaperChange*gc_iCycleTime_Plc;
	IF rTaperCur<rTaperTar THEN
		rTaperCur:=rTaperCur+rDeltTaper;
		IF rTaperCur>=rTaperTar THEN
			rTaperCur:=rTaperTar;
		END_IF
	ELSIF rTaperCur>rTaperTar THEN
		rTaperCur:=rTaperCur-rDeltTaper;
		IF rTaperCur<=rTaperTar THEN
			rTaperCur:=rTaperTar;
		END_IF
	ELSE;
	END_IF
	pstStGrpParam^.lrTaper_Cur_Uw:=rTaperCur;
	(*放牵*)
	rTaperTar:=pstStGrpParam^.lrTaper_Begin_If;
	rTaperCur:=pstStGrpParam^.lrTaper_Cur_If;
	rDeltTaper:=rMaxTaper/iTimeTaperChange*gc_iCycleTime_Plc;
	IF rTaperCur<rTaperTar THEN
		rTaperCur:=rTaperCur+rDeltTaper;
		IF rTaperCur>=rTaperTar THEN
			rTaperCur:=rTaperTar;
		END_IF
	ELSIF rTaperCur>rTaperTar THEN
		rTaperCur:=rTaperCur-rDeltTaper;
		IF rTaperCur<=rTaperTar THEN
			rTaperCur:=rTaperTar;
		END_IF
	ELSE;
	END_IF
	pstStGrpParam^.lrTaper_Cur_If:=rTaperCur;
	(*收牵*)
	rTaperTar:=pstStGrpParam^.lrTaper_Begin_Of;
	rTaperCur:=pstStGrpParam^.lrTaper_Cur_Of;
	rDeltTaper:=rMaxTaper/iTimeTaperChange*gc_iCycleTime_Plc;
	IF rTaperCur<rTaperTar THEN
		rTaperCur:=rTaperCur+rDeltTaper;
		IF rTaperCur>=rTaperTar THEN
			rTaperCur:=rTaperTar;
		END_IF
	ELSIF rTaperCur>rTaperTar THEN
		rTaperCur:=rTaperCur-rDeltTaper;
		IF rTaperCur<=rTaperTar THEN
			rTaperCur:=rTaperTar;
		END_IF
	ELSE;
	END_IF
	pstStGrpParam^.lrTaper_Cur_Of:=rTaperCur;
END_IF

(* ---- KS_FB_TaperUnitDeal.st ---- *)
(*@CES
Name=KS_FB_TaperUnitDeal
Type=FunctionBlock
TypeGuid=6f9dac99-8de1-4efc-8465-68ac443b7d08
Guid=440da615-589b-45d5-ab61-0644875fc808
HasDeclaration=True
HasImplementation=True
*)
{DECLARATION}
FUNCTION_BLOCK KS_FB_TaperUnitDeal(*锥度单位处理*)
(*调整不同单位张力最大值的切换代码执行位置|2022.10.16.105041*)
(*2025.1.15.152035 计算收料停机锥度显示值*)
VAR_INPUT
	i_xEn: BOOL;
END_VAR
VAR_OUTPUT
END_VAR
VAR_IN_OUT
	io_byTaperUnitType:BYTE;(*张力单位切换标志|.0 放牵\.1收牵\.2放料\.3收料*)
	io_byTaperUnit_If: BYTE;
	io_byTaperUnit_Of: BYTE;
	io_byTaperUnit_Uw: BYTE;
	io_byTaperUnit_Rw: BYTE;
	io_byTaperUnitConfirm_Uw : BYTE;

END_VAR
VAR
	byLastUnit_Uw: BYTE:=3;(*初始化给一个不一样的值|用于触发开机取初值*)
	byLastUnit_Rw: BYTE:=3;(*初始化给一个不一样的值|用于触发开机取初值*)
	byLastUnit_If: BYTE:=3;(*初始化给一个不一样的值|用于触发开机取初值*)
	byLastUnit_Of: BYTE:=3;(*初始化给一个不一样的值|用于触发开机取初值*)
END_VAR
{IMPLEMENTATION}
IF i_xEn THEN;
ELSE
	RETURN;
END_IF

(**处理单位切换标志*)
IF io_byTaperUnitType<>0 THEN
	IF io_byTaperUnitType.0 THEN(*放牵切换*)
		io_byTaperUnit_If:=io_byTaperUnit_If+1;
		IF io_byTaperUnit_If>2 THEN
			io_byTaperUnit_If:=0;
		END_IF
	ELSIF io_byTaperUnitType.1 THEN(*收牵切换*)
		io_byTaperUnit_Of:=io_byTaperUnit_Of+1;
		IF io_byTaperUnit_Of>2 THEN
			io_byTaperUnit_Of:=0;
		END_IF
	ELSIF io_byTaperUnitType.2 THEN(*放料切换*)
		io_byTaperUnit_Uw:=io_byTaperUnit_Uw+1;
		IF io_byTaperUnit_Uw>2 THEN
			io_byTaperUnit_Uw:=0;
		END_IF
	ELSIF io_byTaperUnitType.3 THEN(*收料切换*)
		io_byTaperUnit_Rw:=io_byTaperUnit_Rw+1;
		IF io_byTaperUnit_Rw>2 THEN
			io_byTaperUnit_Rw:=0;
		END_IF
	ELSE;
	END_IF
	(*清除单位切换按钮*)
	io_byTaperUnitType:=0;
END_IF

(*放料处理*)
(*
g_rTaperMax_Uw:=100;
IF io_byTaperUnit_Uw=1 THEN(*放料单位|N*)
	g_rTaperMax_Uw:=500;
ELSIF io_byTaperUnit_Uw=2 THEN(*放料单位|Mpa*)
	g_rTaperMax_Uw:=1;
END_IF
*)
KS_CovertUnit_Taper(
	ADR(io_byTaperUnit_Uw)(*i_pbyUnit*),
	i_pstStGrpParam^.byTaperUnitConfirm_Uw.0(*i_xConfirmN*),
	i_pstStGrpParam^.byTaperUnitConfirm_Uw.1(*i_xConfirmMpa*),
	ADR(i_pstStGrpParam^.rPercentMatchN_Uw)(*i_prConfirmTaperPercentMatchN*),
	ADR(i_pstStGrpParam^.rPercentMatchMpa_Uw)(*i_prConfirmTaperPercentMatchMpa*),
	i_pstStGrpParam^.rN_Uw(*i_rConfirmTaperN*),
	i_pstStGrpParam^.rMpa_Uw(*i_rConfirmTaperMpa*),
	ADR(i_pstStGrpParam^.rTaperValueBegin_Hmi_Uw)(*i_prTaperValueBegin_Hmi*),
	ADR(i_pstStGrpParam^.rTaperValueEnd_Hmi_Uw)(*i_prTaperValueEnd_Hmi*),
	ADR(i_pstStGrpParam^.rTaperValueCur_Hmi_Uw)(*i_prTaperValueCur_Hmi*),

	ADR(byLastUnit_Uw)(*i_pbyLastUnit*),
	ADR(i_pstStGrpParam^.lrTaper_Begin_Uw)(*i_plrTaperPencent_Begin*),
	ADR(i_pstStGrpParam^.lrTaper_End_Uw)(*i_plrTaperPencent_End*),
	i_pstStGrpParam^.lrTaper_Cur_Uw(*i_lrTaperPencent_Cur*),
	(*2025.1.15.153326+*)
	0(*i_pbyInitTaper*),
	0(*i_prInitTaper_Hmi*));
(*2022.10.16.104937*)
g_rTaperMax_Uw:=100;
IF io_byTaperUnit_Uw=1 THEN(*放料单位|N*)
	g_rTaperMax_Uw:=500;
ELSIF io_byTaperUnit_Uw=2 THEN(*放料单位|Mpa*)
	g_rTaperMax_Uw:=1;
END_IF
(*清除确认按钮*)
i_pstStGrpParam^.byTaperUnitConfirm_Uw:=0;

(*收料处理*)
(*
g_rTaperMax_Rw:=100;
IF io_byTaperUnit_Rw=1 THEN(*放料单位|N*)
	g_rTaperMax_Rw:=500;
ELSIF io_byTaperUnit_Rw=2 THEN(*放料单位|Mpa*)
	g_rTaperMax_Rw:=1;
END_IF
*)
KS_CovertUnit_Taper(
	ADR(io_byTaperUnit_Rw)(*i_pbyUnit*),
	i_pstStGrpParam^.byTaperUnitConfirm_Rw.0(*i_xConfirmN*),
	i_pstStGrpParam^.byTaperUnitConfirm_Rw.1(*i_xConfirmMpa*),
	ADR(i_pstStGrpParam^.rPercentMatchN_Rw)(*i_prConfirmTaperPercentMatchN*),
	ADR(i_pstStGrpParam^.rPercentMatchMpa_Rw)(*i_prConfirmTaperPercentMatchMpa*),
	i_pstStGrpParam^.rN_Rw(*i_rConfirmTaperN*),
	i_pstStGrpParam^.rMpa_Rw(*i_rConfirmTaperMpa*),
	ADR(i_pstStGrpParam^.rTaperValueBegin_Hmi_Rw)(*i_prTaperValueBegin_Hmi*),
	ADR(i_pstStGrpParam^.rTaperValueEnd_Hmi_Rw)(*i_prTaperValueEnd_Hmi*),
	ADR(i_pstStGrpParam^.rTaperValueCur_Hmi_Rw)(*i_prTaperValueCur_Hmi*),
	ADR(byLastUnit_Rw)(*i_pbyLastUnit*),
	ADR(i_pstStGrpParam^.lrTaper_Begin_Rw)(*i_plrTaperPencent_Begin*),
	ADR(i_pstStGrpParam^.lrTaper_End_Rw)(*i_plrTaperPencent_End*),
	i_pstStGrpParam^.lrTaper_Cur_Rw(*i_lrTaperPencent_Cur*),
	(*2025.1.15.153326+*)
	ADR(i_pstStGrpParam^.byInitTaper_Rw)(*i_pbyInitTaper*),
	ADR(i_pstStGrpParam^.rInitTaper_Hmi_Rw)(*i_prInitTaper_Hmi*));
(*2022.10.16.104955*)
g_rTaperMax_Rw:=100;
IF io_byTaperUnit_Rw=1 THEN(*放料单位|N*)
	g_rTaperMax_Rw:=500;
ELSIF io_byTaperUnit_Rw=2 THEN(*放料单位|Mpa*)
	g_rTaperMax_Rw:=1;
END_IF
(*清除确认按钮*)
i_pstStGrpParam^.byTaperUnitConfirm_Rw:=0;

(*放牵处理*)
(*
g_rTaperMax_If:=100;
IF io_byTaperUnit_If=1 THEN(*放料单位|N*)
	g_rTaperMax_If:=500;
ELSIF io_byTaperUnit_If=2 THEN(*放料单位|Mpa*)
	g_rTaperMax_If:=1;
END_IF
*)
KS_CovertUnit_Taper(
	ADR(io_byTaperUnit_If)(*i_pbyUnit*),
	i_pstStGrpParam^.byTaperUnitConfirm_If.0(*i_xConfirmN*),
	i_pstStGrpParam^.byTaperUnitConfirm_If.1(*i_xConfirmMpa*),
	ADR(i_pstStGrpParam^.rPercentMatchN_If)(*i_prConfirmTaperPercentMatchN*),
	ADR(i_pstStGrpParam^.rPercentMatchMpa_If)(*i_prConfirmTaperPercentMatchMpa*),
	i_pstStGrpParam^.rN_If(*i_rConfirmTaperN*),
	i_pstStGrpParam^.rMpa_If(*i_rConfirmTaperMpa*),
	ADR(i_pstStGrpParam^.rTaperValueBegin_Hmi_If)(*i_prTaperValueBegin_Hmi*),
	ADR(i_pstStGrpParam^.rTaperValueEnd_Hmi_If)(*i_prTaperValueEnd_Hmi*),
	ADR(i_pstStGrpParam^.rTaperValueCur_Hmi_If)(*i_prTaperValueCur_Hmi*),
	ADR(byLastUnit_If)(*i_pbyLastUnit*),
	ADR(i_pstStGrpParam^.lrTaper_Begin_If)(*i_plrTaperPencent_Begin*),
	ADR(i_pstStGrpParam^.lrTaper_End_If)(*i_plrTaperPencent_End*),
	i_pstStGrpParam^.lrTaper_Cur_If(*i_lrTaperPencent_Cur*),
	(*2025.1.15.153326+*)
	0(*i_pbyInitTaper*),
	0(*i_prInitTaper_Hmi*));
(*2022.10.16.105013*)
g_rTaperMax_If:=100;
IF io_byTaperUnit_If=1 THEN(*放料单位|N*)
	g_rTaperMax_If:=500;
ELSIF io_byTaperUnit_If=2 THEN(*放料单位|Mpa*)
	g_rTaperMax_If:=1;
END_IF
(*清除确认按钮*)
i_pstStGrpParam^.byTaperUnitConfirm_If:=0;

(*收牵处理*)
(*
g_rTaperMax_of:=100;
IF io_byTaperUnit_Of=1 THEN(*放料单位|N*)
	g_rTaperMax_of:=500;
ELSIF io_byTaperUnit_Of=2 THEN(*放料单位|Mpa*)
	g_rTaperMax_of:=1;
END_IF
*)
KS_CovertUnit_Taper(
	ADR(io_byTaperUnit_Of)(*i_pbyUnit*),
	i_pstStGrpParam^.byTaperUnitConfirm_Of.0(*i_xConfirmN*),
	i_pstStGrpParam^.byTaperUnitConfirm_Of.1(*i_xConfirmMpa*),
	ADR(i_pstStGrpParam^.rPercentMatchN_Of)(*i_prConfirmTaperPercentMatchN*),
	ADR(i_pstStGrpParam^.rPercentMatchMpa_Of)(*i_prConfirmTaperPercentMatchMpa*),
	i_pstStGrpParam^.rN_Of(*i_rConfirmTaperN*),
	i_pstStGrpParam^.rMpa_Of(*i_rConfirmTaperMpa*),
	ADR(i_pstStGrpParam^.rTaperValueBegin_Hmi_Of)(*i_prTaperValueBegin_Hmi*),
	ADR(i_pstStGrpParam^.rTaperValueEnd_Hmi_Of)(*i_prTaperValueEnd_Hmi*),
	ADR(i_pstStGrpParam^.rTaperValueCur_Hmi_Of)(*i_prTaperValueCur_Hmi*),
	ADR(byLastUnit_Of)(*i_pbyLastUnit*),
	ADR(i_pstStGrpParam^.lrTaper_Begin_Of)(*i_plrTaperPencent_Begin*),
	ADR(i_pstStGrpParam^.lrTaper_End_Of)(*i_plrTaperPencent_End*),
	i_pstStGrpParam^.lrTaper_Cur_Of(*i_lrTaperPencent_Cur*),
	(*2025.1.15.153326+*)
	0(*i_pbyInitTaper*),
	0(*i_prInitTaper_Hmi*));
(*2022.10.16.105028*)
g_rTaperMax_of:=100;
IF io_byTaperUnit_Of=1 THEN(*放料单位|N*)
	g_rTaperMax_of:=500;
ELSIF io_byTaperUnit_Of=2 THEN(*放料单位|Mpa*)
	g_rTaperMax_of:=1;
END_IF
(*清除确认按钮*)
i_pstStGrpParam^.byTaperUnitConfirm_Of:=0;

(* ---- KS_FB_TaperUnitDeal_New.st ---- *)
(*@CES
Name=KS_FB_TaperUnitDeal_New
Type=FunctionBlock
TypeGuid=6f9dac99-8de1-4efc-8465-68ac443b7d08
Guid=029751e0-fe3d-4f68-a3f4-ab7fe94fc43b
HasDeclaration=True
HasImplementation=True
*)
{DECLARATION}
FUNCTION_BLOCK KS_FB_TaperUnitDeal_New(*锥度单位处理*)
(*调整不同单位张力最大值的切换代码执行位置|2022.10.16.105041*)
(*2025.1.15.152035 计算收料停机锥度显示值*)
VAR_INPUT
	i_xEn: BOOL;
	i_rN: REAL;
	i_rMpa: REAL;
	i_pbyInitTaper: POINTER TO BYTE;
	i_prInitTaper_Hmi: POINTER TO REAL;
END_VAR
VAR_OUTPUT
END_VAR
VAR_IN_OUT
	io_xTaperUnitType:BOOL;(*张力单位切换标志|.0 放牵\.1收牵\.2放料\.3收料*)
	io_byTaperUnit: BYTE;
	io_byTaperUnitConfirm : BYTE;
	io_rPercentMatchN: REAL;
	io_rPercentMatchMpa: REAL;
	io_rTaperValueBegin_Hmi: REAL;
	io_rTaperValueEnd_Hmi: REAL;
	io_rTaperValueCur_Hmi: REAL;
	io_rTaper_Begin: REAL;
	io_rTaper_End: REAL;
	io_rTaper_Cur: REAL;
	io_rTaperMax: REAL;

END_VAR
VAR
	byLastUnit: BYTE:=3;(*初始化给一个不一样的值|用于触发开机取初值*)
END_VAR
{IMPLEMENTATION}
IF i_xEn THEN;
ELSE
	RETURN;
END_IF

(**处理单位切换标志*)
IF io_xTaperUnitType THEN(*放牵切换*)
	io_byTaperUnit:=io_byTaperUnit+1;
	IF io_byTaperUnit>2 THEN
		io_byTaperUnit:=0;
	END_IF

ELSE;
END_IF
(*清除单位切换按钮*)
io_xTaperUnitType:=FALSE;

KS_CovertUnit_Taper(
	ADR(io_byTaperUnit)(*i_pbyUnit*),
	io_byTaperUnitConfirm.0(*i_xConfirmN*),
	io_byTaperUnitConfirm.1(*i_xConfirmMpa*),
	ADR(io_rPercentMatchN)(*i_prConfirmTaperPercentMatchN*),
	ADR(io_rPercentMatchMpa)(*i_prConfirmTaperPercentMatchMpa*),
	i_rN(*i_rConfirmTaperN*),
	i_rMpa(*i_rConfirmTaperMpa*),
	ADR(io_rTaperValueBegin_Hmi)(*i_prTaperValueBegin_Hmi*),
	ADR(io_rTaperValueEnd_Hmi)(*i_prTaperValueEnd_Hmi*),
	ADR(io_rTaperValueCur_Hmi)(*i_prTaperValueCur_Hmi*),

	ADR(byLastUnit)(*i_pbyLastUnit*),
	ADR(io_rTaper_Begin)(*i_plrTaperPencent_Begin*),
	ADR(io_rTaper_End)(*i_plrTaperPencent_End*),
	io_rTaper_Cur(*i_lrTaperPencent_Cur*),
	(*2025.1.15.153326+*)
	i_pbyInitTaper,
	i_prInitTaper_Hmi);
(*2022.10.16.104937*)
io_rTaperMax:=100;
IF io_byTaperUnit=1 THEN(*放料单位|N*)
	io_rTaperMax:=500;
ELSIF io_byTaperUnit=2 THEN(*放料单位|Mpa*)
	io_rTaperMax:=1;
END_IF
(*清除确认按钮*)
io_byTaperUnitConfirm:=0;
